Fanuc KAREL source: ko00066.KL

PROGRAM KO00066
%STACKSIZE=65535
%PRIORITY=65535
%NOLOCKGROUP
VAR
P1 : XYZWPREXT
P2 : POSITION
F : BOOLEAN
OUT : XYZWPR
BEGIN
F=TRUE
OUT=MIRROR(P1,P2,F)
END KO00066
